Fanuc KAREL source: KB00004.KL

PROGRAM KB00004
%NOLOCKGROUP
VAR
BEGIN
  ACT_SCREEN
END KB00004
